// TIA Portal V20 export
// export: Created 2026-10-12T05:35:22.2104437Z, ExportSetting WithDefaults, DisplayName Totally Integrated Automation Portal, DisplayVersion V20, DisplayName TIA Portal Openness, DisplayVersion V20, DisplayName TIA Portal Teamcenter Gateway, DisplayVersion V20, DisplayName TIA Portal Version Control Interface, DisplayVersion V20, DisplayName SINAMICS Startdrive Advanced, DisplayVersion V20 SP1 Update 2, DisplayName SINAMICS Startdrive G110M, G120, G120C, G120D, G120P, G115D, DisplayVersion V20 SP1 Update 2, DisplayName SINAMICS Startdrive G130, G150, S120, S150, SINAMICS MV, G220, S200, S210, DisplayVersion V20 SP1 Update 2, DisplayName STEP 7 Professional, DisplayVersion V20, DisplayName STEP 7 Safety, DisplayVersion V20, DisplayName WinCC Basic/Comfort/Advanced, DisplayVersion V20, DisplayName WinCC Professional, DisplayVersion V20, DisplayName WinCC Unified, DisplayVersion V20
FUNCTION "FRK_ClockTick" : Void   // FC4, SCL
{ S7_Optimized_Access := 'TRUE' }
VERSION : 0.1
// Shared command kernel v0.1. Core 2.2 / 6.1 / 3.14 / 8.11.
//  Generated enum/rationalization values come from Core authorities.
// stored: AutoNumber true, IsIECCheckEnabled false, SetENOAutomatically false, UDAEnableTagReadback false
   VAR_TEMP
      DeltaS : LReal;
   END_VAR
BEGIN

   #DeltaS := RUNTIME("FRK_Clock".Mem);
   IF #DeltaS < 0.0 OR #DeltaS > 60.0 THEN
       #DeltaS := 0.0;
   END_IF;
   "FRK_Clock".AccMs := "FRK_Clock".AccMs + #DeltaS * 1000.0;
   IF "FRK_Clock".AccMs >= 4294967296.0 THEN
       "FRK_Clock".AccMs := "FRK_Clock".AccMs - 4294967296.0;
   END_IF;
   "FRK_Clock".NowMs := TRUNC_UDINT("FRK_Clock".AccMs);
END_FUNCTION
